PROGRAM Control_FBD
VAR
	
	batLevel1 : BOOL;
	batLevel2: BOOL;
	batLevel3: BOOL;
	
	mxRun : BOOL;
	qxMotorUp : BOOL;
	qxMotorDown: BOOL;
	
	SR1: SR;
	RS1: RS;
	TOF_1: TOF;
	TON_1: TON;
END_VAR
VAR // added by the converter: edge detectors and wires of the graphical bodies
    _w1, _w2, _w3 : BOOL;
END_VAR

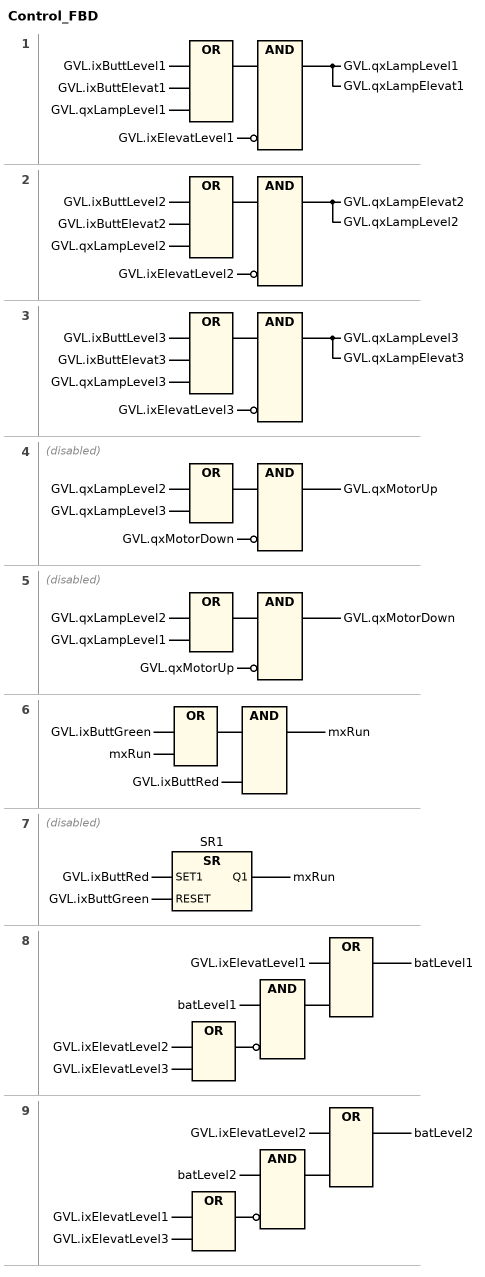
// NETWORK 1
_w1 := (GVL.ixButtLevel1 OR GVL.ixButtElevat1 OR GVL.qxLampLevel1) AND NOT GVL.ixElevatLevel1;
GVL.qxLampLevel1 := _w1;
GVL.qxLampElevat1 := _w1;

// NETWORK 2
_w2 := (GVL.ixButtLevel2 OR GVL.ixButtElevat2 OR GVL.qxLampLevel2) AND NOT GVL.ixElevatLevel2;
GVL.qxLampElevat2 := _w2;
GVL.qxLampLevel2 := _w2;

// NETWORK 3
_w3 := (GVL.ixButtLevel3 OR GVL.ixButtElevat3 OR GVL.qxLampLevel3) AND NOT GVL.ixElevatLevel3;
GVL.qxLampLevel3 := _w3;
GVL.qxLampElevat3 := _w3;

// NETWORK 4 (disabled)
// GVL.qxMotorUp := (GVL.qxLampLevel2 OR GVL.qxLampLevel3) AND NOT GVL.qxMotorDown;

// NETWORK 5 (disabled)
// GVL.qxMotorDown := (GVL.qxLampLevel2 OR GVL.qxLampLevel1) AND NOT GVL.qxMotorUp;

// NETWORK 6
mxRun := (GVL.ixButtGreen OR mxRun) AND GVL.ixButtRed;

// NETWORK 7 (disabled)
// SR1(SET1 := GVL.ixButtRed, RESET := GVL.ixButtGreen); // SR
// mxRun := SR1.Q1;

// NETWORK 8
batLevel1 := GVL.ixElevatLevel1 OR batLevel1 AND NOT (GVL.ixElevatLevel2 OR GVL.ixElevatLevel3);

// NETWORK 9
batLevel2 := GVL.ixElevatLevel2 OR batLevel2 AND NOT (GVL.ixElevatLevel1 OR GVL.ixElevatLevel3);

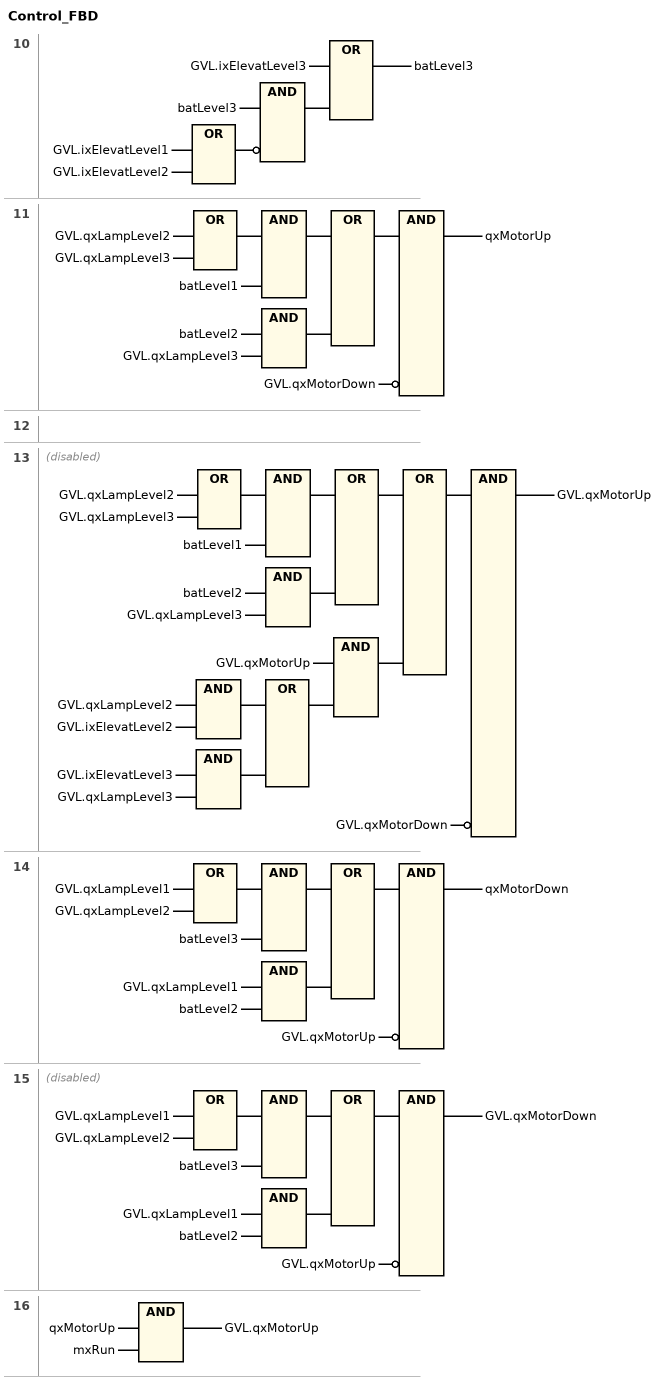
// NETWORK 10
batLevel3 := GVL.ixElevatLevel3 OR batLevel3 AND NOT (GVL.ixElevatLevel1 OR GVL.ixElevatLevel2);

// NETWORK 11
qxMotorUp := ((GVL.qxLampLevel2 OR GVL.qxLampLevel3) AND batLevel1 OR batLevel2 AND GVL.qxLampLevel3) AND NOT GVL.qxMotorDown;

// NETWORK 12

// NETWORK 13 (disabled)
// GVL.qxMotorUp := (((GVL.qxLampLevel2 OR GVL.qxLampLevel3) AND batLevel1 OR batLevel2 AND GVL.qxLampLevel3) OR GVL.qxMotorUp AND (GVL.qxLampLevel2 AND GVL.ixElevatLevel2 OR GVL.ixElevatLevel3 AND GVL.qxLampLevel3)) AND NOT GVL.qxMotorDown;

// NETWORK 14
qxMotorDown := ((GVL.qxLampLevel1 OR GVL.qxLampLevel2) AND batLevel3 OR GVL.qxLampLevel1 AND batLevel2) AND NOT GVL.qxMotorUp;

// NETWORK 15 (disabled)
// GVL.qxMotorDown := ((GVL.qxLampLevel1 OR GVL.qxLampLevel2) AND batLevel3 OR GVL.qxLampLevel1 AND batLevel2) AND NOT GVL.qxMotorUp;

// NETWORK 16
GVL.qxMotorUp := qxMotorUp AND mxRun;

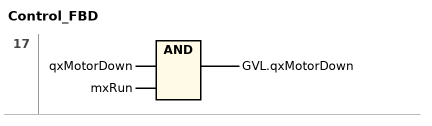
// NETWORK 17
GVL.qxMotorDown := qxMotorDown AND mxRun;

END_PROGRAM

(* stored: Version 1.1.0.1
   POU Control_FBD: Id {912119c4-f197-4ac1-96d5-56b57bc2b241}, SpecialFunc None *)
